VAR_GLOBAL
    bButton AT %I* : BOOL;
    bLightRelay AT %Q* : BOOL;
END_VAR

(* stored: Version 1.1.0.1
   GVL GVL_WorkshopIO: Id {25c89f3f-8e8e-413a-98e1-365895cc7aa8} *)
